(* IEC 61131-3 sources: plc-vscode/tests/st/all/trust-platform/crates/trust-runtime/tests/fixtures/oscat/core/src/23_control_modules, 1 file *)

(* ---- tests.st ---- *)
TEST_PROGRAM oscat_control_modules_basic_helpers_behave
ASSERT_EQUAL(EXPECTED := BYTE#0, ACTUAL := BAND_B(X := BYTE#2, B := BYTE#5));
ASSERT_EQUAL(EXPECTED := BYTE#250, ACTUAL := BAND_B(X := BYTE#250, B := BYTE#5));
ASSERT_NEAR(EXPECTED := REAL#7.0, ACTUAL := CTRL_IN(SET_POINT := REAL#10.0, ACTUAL := REAL#2.0, NOISE := REAL#1.0), DELTA := REAL#0.001);
ASSERT_NEAR(EXPECTED := REAL#4.0, ACTUAL := DEAD_BAND(X := REAL#5.0, L := REAL#1.0), DELTA := REAL#0.001);
ASSERT_NEAR(EXPECTED := REAL#5.0, ACTUAL := DEAD_ZONE(X := REAL#5.0, L := REAL#1.0), DELTA := REAL#0.001);
ASSERT_NEAR(EXPECTED := REAL#0.0, ACTUAL := DEAD_ZONE(X := REAL#0.5, L := REAL#1.0), DELTA := REAL#0.001);
END_TEST_PROGRAM

TEST_PROGRAM oscat_control_modules_control_set_helpers_behave
VAR
    Set1 : CONTROL_SET1;
    Set2 : CONTROL_SET2;
END_VAR

Set1(Kt := REAL#10.0, Tt := REAL#20.0, PI := FALSE, PID := TRUE);
ASSERT_NEAR(EXPECTED := REAL#6.0, ACTUAL := Set1.KP, DELTA := REAL#0.001);
ASSERT_NEAR(EXPECTED := REAL#10.0, ACTUAL := Set1.TN, DELTA := REAL#0.001);
ASSERT_NEAR(EXPECTED := REAL#2.5, ACTUAL := Set1.TV, DELTA := REAL#0.001);
ASSERT_NEAR(EXPECTED := REAL#0.6, ACTUAL := Set1.KI, DELTA := REAL#0.001);
ASSERT_NEAR(EXPECTED := REAL#15.0, ACTUAL := Set1.KD, DELTA := REAL#0.001);

Set2(KS := REAL#2.0, TU := REAL#3.0, TG := REAL#12.0, PI := TRUE, PID := FALSE);
ASSERT_NEAR(EXPECTED := REAL#1.8, ACTUAL := Set2.KP, DELTA := REAL#0.001);
ASSERT_NEAR(EXPECTED := REAL#9.99, ACTUAL := Set2.TN, DELTA := REAL#0.02);
ASSERT_NEAR(EXPECTED := REAL#0.0, ACTUAL := Set2.TV, DELTA := REAL#0.001);
ASSERT_NEAR(EXPECTED := REAL#0.18018, ACTUAL := Set2.KI, DELTA := REAL#0.001);
ASSERT_NEAR(EXPECTED := REAL#0.0, ACTUAL := Set2.KD, DELTA := REAL#0.001);
END_TEST_PROGRAM

TEST_PROGRAM oscat_control_modules_hysteresis_helpers_behave
VAR
    H1 : HYST;
    H2 : HYST_1;
    H3 : HYST_2;
    H4 : HYST_3;
END_VAR

H1(IN := REAL#12.0, HIGH_LIMIT := REAL#10.0, LOW_LIMIT := REAL#8.0);
ASSERT_TRUE(IN := H1.Q);
ASSERT_FALSE(IN := H1.WIN);

H2(IN := REAL#5.0, high := REAL#4.0, low := REAL#2.0);
ASSERT_TRUE(IN := H2.Q);
ASSERT_FALSE(IN := H2.WIN);

H3(IN := REAL#12.0, VAL := REAL#10.0, HYS := REAL#2.0);
ASSERT_TRUE(IN := H3.Q);
ASSERT_FALSE(IN := H3.WIN);

H4(IN := REAL#4.0, hyst := REAL#2.0, val1 := REAL#6.0, val2 := REAL#8.0);
ASSERT_TRUE(IN := H4.Q1);
ASSERT_FALSE(IN := H4.Q2);
END_TEST_PROGRAM

TEST_PROGRAM oscat_control_modules_hyst_2_retains_state_inside_window
VAR
    H3 : HYST_2;
    QHigh : BOOL := FALSE;
    WinHigh : BOOL := FALSE;
    QWindow : BOOL := FALSE;
    WinWindow : BOOL := FALSE;
    QLow : BOOL := FALSE;
    WinLow : BOOL := FALSE;
END_VAR

H3(IN := REAL#12.0, VAL := REAL#10.0, HYS := REAL#2.0);
QHigh := H3.Q;
WinHigh := H3.WIN;

H3(IN := REAL#9.5, VAL := REAL#10.0, HYS := REAL#2.0);
QWindow := H3.Q;
WinWindow := H3.WIN;

H3(IN := REAL#8.5, VAL := REAL#10.0, HYS := REAL#2.0);
QLow := H3.Q;
WinLow := H3.WIN;

ASSERT_TRUE(IN := QHigh);
ASSERT_FALSE(IN := WinHigh);
ASSERT_TRUE(IN := QWindow);
ASSERT_TRUE(IN := WinWindow);
ASSERT_FALSE(IN := QLow);
ASSERT_FALSE(IN := WinLow);
END_TEST_PROGRAM

TEST_PROGRAM oscat_control_modules_ctrl_pid_manual_clamp_behaves
VAR
    Ctrl : CTRL_PID;
END_VAR

Ctrl(
    ACT := REAL#0.0,
    SET_POINT := REAL#10.0,
    SUP := REAL#0.0,
    OFS := REAL#1.0,
    M_I := REAL#50.0,
    MAN := TRUE,
    RST := FALSE,
    KP := REAL#2.0,
    TN := REAL#1.0,
    TV := REAL#0.0,
    LL := REAL#0.0,
    LH := REAL#10.0
);

ASSERT_NEAR(EXPECTED := REAL#10.0, ACTUAL := Ctrl.Y, DELTA := REAL#0.001);
ASSERT_NEAR(EXPECTED := REAL#10.0, ACTUAL := Ctrl.DIFF, DELTA := REAL#0.001);
ASSERT_TRUE(IN := Ctrl.LIM);
END_TEST_PROGRAM

TEST_PROGRAM oscat_control_modules_environmental_functions_behave
VAR
    RhoAir : REAL;
    Condensation : REAL;
END_VAR

ASSERT_TRUE(IN := OSCAT_BASIC_Constants());
ASSERT_NEAR(EXPECTED := REAL#20.0964, ACTUAL := AIR_ENTHALPY(T := REAL#20.0, RH := REAL#0.0), DELTA := REAL#0.01);
ASSERT_NEAR(EXPECTED := REAL#0.0, ACTUAL := DEW_CON(RH := REAL#0.0, T := REAL#20.0), DELTA := REAL#0.0001);
ASSERT_NEAR(EXPECTED := REAL#20.0, ACTUAL := DEW_TEMP(RH := REAL#100.0, T := REAL#20.0), DELTA := REAL#0.01);
Condensation := DEW_CON(RH := REAL#50.0, T := REAL#20.0);
ASSERT_NEAR(EXPECTED := REAL#50.0, ACTUAL := DEW_RH(VC := Condensation, T := REAL#20.0), DELTA := REAL#0.1);
RhoAir := AIR_DENSITY(T := REAL#20.0, P := REAL#101325.0, RH := REAL#50.0);
ASSERT_NEAR(EXPECTED := REAL#1.2, ACTUAL := RhoAir, DELTA := REAL#0.1);
ASSERT_NEAR(EXPECTED := REAL#4.228, ACTUAL := WATER_CP(T := REAL#0.0), DELTA := REAL#0.001);
ASSERT_NEAR(EXPECTED := REAL#42.1, ACTUAL := WATER_ENTHALPY(T := REAL#10.0), DELTA := REAL#0.1);
ASSERT_NEAR(EXPECTED := REAL#1000.0, ACTUAL := WATER_DENSITY(T := REAL#4.0, Sat := FALSE), DELTA := REAL#1.0);
ASSERT_NEAR(EXPECTED := REAL#2.0944, ACTUAL := TANK_VOL2(TR := REAL#1.0, H := REAL#1.0), DELTA := REAL#0.001);
ASSERT_NEAR(EXPECTED := REAL#3.14159, ACTUAL := TANK_VOL1(TR := REAL#1.0, TL := REAL#2.0, H := REAL#1.0), DELTA := REAL#0.01);
ASSERT_NEAR(EXPECTED := REAL#5.0, ACTUAL := WCT(T := REAL#5.0, V := REAL#2.0), DELTA := REAL#0.001);
END_TEST_PROGRAM

TEST_PROGRAM oscat_control_modules_building_blocks_behave
VAR
    Coil : ACTUATOR_COIL;
    Window : TIMER_1;
    BoilerCtrl : BOILER;
    HeatingCurve : HEAT_TEMP;
    OutsideTemp : TEMP_EXT;
END_VAR

Coil(IN := TRUE);
ASSERT_TRUE(IN := Coil.OUT);
ASSERT_EQUAL(EXPECTED := BYTE#101, ACTUAL := Coil.STATUS);

Window(E := TRUE, DTI := DT#2026-01-04-10:30:00, START := TOD#10:00:00, DURATION := T#1h, DAY := BYTE#127);
ASSERT_TRUE(IN := Window.Q);

BoilerCtrl(T_upper := REAL#45.0, T_lower := REAL#45.0, Pressure := TRUE, enable := TRUE, Req_1 := FALSE, Req_2 := FALSE, Boost := FALSE);
ASSERT_TRUE(IN := BoilerCtrl.Heat);
ASSERT_FALSE(IN := BoilerCtrl.error);
ASSERT_EQUAL(EXPECTED := BYTE#102, ACTUAL := BoilerCtrl.status);

HeatingCurve(T_EXT := REAL#0.0, T_INT := REAL#20.0, OFFSET := REAL#0.0, T_REQ := REAL#0.0);
ASSERT_TRUE(IN := HeatingCurve.HEAT);
ASSERT_NEAR(EXPECTED := REAL#52.4, ACTUAL := HeatingCurve.TY, DELTA := REAL#2.0);

OutsideTemp(t_ext1 := REAL#-15.0, t_ext2 := REAL#-14.0, t_ext3 := REAL#-16.0, t_ext_config := BYTE#0, dt_in := DT#2026-01-15-12:00:00);
ASSERT_TRUE(IN := OutsideTemp.heat);
ASSERT_FALSE(IN := OutsideTemp.cool);
END_TEST_PROGRAM
